{attribute 'qualified_only'}
{attribute 'strict'}
{attribute 'to_string'}
TYPE E_INSTANCE_CHECK :
(
  NULL,

	POINTER_COLLECTOR_ITF_INVALID := 9000,
  INVALID_INSTANCE_CONTROL_REFERENCE,
  INVALID_INSTANCE_STATE_REFERENCE,
  PROCESS_ID_ZERO := 9100,
  PROCESS_ID_MAX  := 9200,
  PROCESS_ID_NOTEQUAL_COLLECTOR_ID := 9300,
  PROCESS_LIST_ITF_INDEX_INVALID := 9400,
  TICKET_LIST_ITF_INVALID,

  CTRL_CYCLIC_LIST_REFERENCE_INVALID  := 9500,
  STATE_CYCLIC_LIST_REFERENCE_INVALID,
  DATA_CYCLIC_LIST_REFERENCE_INVALID,
  

  CHECK_DONE := 10000
)UINT;
END_TYPE

(* stored: Version 1.1.0.1
   DUT E_INSTANCE_CHECK: Id {928a9ea8-18df-4fd8-9d64-30e0e715bb30} *)
